{region 'Documentation'}
(*!
<summary>Character codes use WORD; exact comparison without a mask.</summary>
<description>

Searches the selected IN range for the complete contiguous Expected pattern.

StartIndex is an absolute declared IN index, not an offset. Length selects 1..255
elements; the complete selected range must fit IN. Invalid references or ranges report
Error.

Keep supplied arrays stable for the call. Input data is read, not copied or retained as a
snapshot.

The complete Expected pattern must be nonempty and fit the selected IN range; an
oversized pattern reports Error, not a missing-match result.

</description>
*)
{endregion}
FUNCTION_BLOCK AssertArrayContainsArray_WChar EXTENDS AssertionBase
VAR_INPUT
    StartIndex : DINT; //! First selected index in IN; uses the array's declared index range, not a zero-based offset.
    Length : USINT; //! Number of searched elements, from 1 through 255.
END_VAR
VAR_IN_OUT CONSTANT
    IN : ARRAY[*] OF WORD; //! Read-only search data; keep stable during the call.
    Expected : ARRAY[*] OF WORD; //! Read-only expected sequence starting at its own lower bound; must fit the selected actual range.
END_VAR

SUPER^();

{region 'Documentation'}
(*!
<summary>Validate configuration before searching the selected range.</summary>
*)
{endregion}
METHOD PROTECTED Assert
VAR
    InLowerIndex : DINT;
    InUpperIndex : DINT;
    EndIndex : LINT;
    Offset : LINT;
    InIndex : DINT;
    ExpectedLowerIndex : DINT;
    ExpectedUpperIndex : DINT;
    ExpectedLength : LINT;
    ExpectedIndex : DINT;
    CandidateOffset : LINT;
    PatternFound : BOOL;
    PatternMatches : BOOL;
    Message : STRING(GVL_Constants.MessageLength);
END_VAR
IF NOT EvaluationActive THEN
    RETURN;
END_IF;

IF Result = E_Result.Error THEN
    RETURN;
END_IF;

// C0371: FB input is checked here before any reference access.
{warning disable C0371}
IF NOT __ISVALIDREF(IN) THEN
    Error(Message := 'Assertion error: IN reference is invalid.');
    RETURN;
END_IF;

IF NOT __ISVALIDREF(Expected) THEN
    Error(Message := 'Assertion error: Expected reference is invalid.');
    RETURN;
END_IF;

InLowerIndex := LOWER_BOUND(IN, 1);
InUpperIndex := UPPER_BOUND(IN, 1);
EndIndex := DINT_TO_LINT(StartIndex) + USINT_TO_LINT(Length) - 1;

ExpectedLowerIndex := LOWER_BOUND(Expected, 1);
ExpectedUpperIndex := UPPER_BOUND(Expected, 1);
ExpectedLength := DINT_TO_LINT(ExpectedUpperIndex) - DINT_TO_LINT(ExpectedLowerIndex) + 1;

IF (Length = 0)
    OR (ExpectedLength <= 0) OR (ExpectedLength > USINT_TO_LINT(Length))
    OR (StartIndex < InLowerIndex) OR (StartIndex > InUpperIndex)
    OR (EndIndex > DINT_TO_LINT(InUpperIndex)) THEN
    Message := CONCAT('Assertion error: array range or pattern is invalid. StartIndex = ',
        DINT_TO_STRING(StartIndex));
    Message := CONCAT(Message, ', Length = ');
    Message := CONCAT(Message, USINT_TO_STRING(Length));
    Message := CONCAT(Message, ', ExpectedLength = ');
    Message := CONCAT(Message, LINT_TO_STRING(ExpectedLength));
    Message := CONCAT(Message, '.');
    Error(Message := Message);
    RETURN;
END_IF;

IF Result = E_Result.Failed THEN
    RETURN;
END_IF;

PatternFound := FALSE;
FOR CandidateOffset := 0 TO USINT_TO_LINT(Length) - ExpectedLength DO
    PatternMatches := TRUE;
    FOR Offset := 0 TO ExpectedLength - 1 DO
        InIndex := LINT_TO_DINT(DINT_TO_LINT(StartIndex) + CandidateOffset + Offset);
        ExpectedIndex := LINT_TO_DINT(DINT_TO_LINT(ExpectedLowerIndex) + Offset);
        IF IN[InIndex] <> Expected[ExpectedIndex] THEN
            PatternMatches := FALSE;
            EXIT;
        END_IF;
    END_FOR;

    IF PatternMatches THEN
        PatternFound := TRUE;
        EXIT;
    END_IF;
END_FOR;

IF NOT PatternFound THEN
    Message := CONCAT('Assertion failed: array range does not contain Expected pattern. ExpectedRange = [',
        DINT_TO_STRING(ExpectedLowerIndex));
    Message := CONCAT(Message, '..');
    Message := CONCAT(Message, DINT_TO_STRING(ExpectedUpperIndex));
    Message := CONCAT(Message, '], ActualRange = [');
    Message := CONCAT(Message, DINT_TO_STRING(StartIndex));
    Message := CONCAT(Message, '..');
    Message := CONCAT(Message, LINT_TO_STRING(EndIndex));
    Message := CONCAT(Message, ']');
    Message := CONCAT(Message, '.');
    Fail(Message := Message);
    RETURN;
END_IF;

Pass();
{warning restore C0371}
END_METHOD

END_FUNCTION_BLOCK

(* stored: Version 1.1.0.1
   POU AssertArrayContainsArray_WChar: Id {70fb1c2f-2339-4b98-9f50-f180fc08f24c}, SpecialFunc None
   Folder Internal: Id {a74caa15-a3c8-4f49-9af8-4df6f7942b8c}
   Method Assert: Id {9fee300e-8ebe-416f-a16d-3461f5893f5b} *)
